Fanuc KAREL source: NC0010.KL

PROGRAM NC0010
%NOLOCKGROUP
ROUTINE R
VAR
  X : INTEGER
BEGIN
  X = 1
  IF X = 1 THEN
    IF X = 1 THEN
      IF X = 1 THEN
        IF X = 1 THEN
          IF X = 1 THEN
            IF X = 1 THEN
              IF X = 1 THEN
                IF X = 1 THEN
                  IF X = 1 THEN
                    IF X = 1 THEN
                      IF X = 1 THEN
                        IF X = 1 THEN
                          IF X = 1 THEN
                            IF X = 1 THEN
                              IF X = 1 THEN
                                IF X = 1 THEN
                                  IF X = 1 THEN
                                    IF X = 1 THEN
                                      X = X + 1
                                    ELSE
                                      X = X + 2
                                    ENDIF
                                  ELSE
                                    X = X + 2
                                  ENDIF
                                ELSE
                                  X = X + 2
                                ENDIF
                              ELSE
                                X = X + 2
                              ENDIF
                            ELSE
                              X = X + 2
                            ENDIF
                          ELSE
                            X = X + 2
                          ENDIF
                        ELSE
                          X = X + 2
                        ENDIF
                      ELSE
                        X = X + 2
                      ENDIF
                    ELSE
                      X = X + 2
                    ENDIF
                  ELSE
                    X = X + 2
                  ENDIF
                ELSE
                  X = X + 2
                ENDIF
              ELSE
                X = X + 2
              ENDIF
            ELSE
              X = X + 2
            ENDIF
          ELSE
            X = X + 2
          ENDIF
        ELSE
          X = X + 2
        ENDIF
      ELSE
        X = X + 2
      ENDIF
    ELSE
      X = X + 2
    ENDIF
  ELSE
    X = X + 2
  ENDIF
END R
BEGIN
  R
END NC0010
